FUNCTION_BLOCK Actuator2OpBaseExt (* Composite Function Block Type *)
  (* Standard: 61499-2 *)
  (* Version 1.0.1, 9/20/2023, ApplicationLibDevTeam, Schneider Electric, First Version *)
  PACKAGE Flexbridge.FestoMPS400;
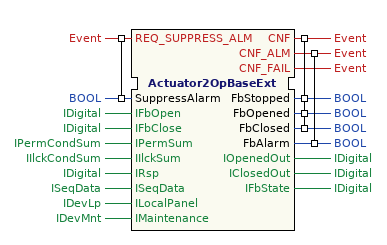
  EVENT_INPUT
    REQ_SUPPRESS_ALM WITH SuppressAlarm; (* Request to update the alarm suppress status *)
  END_EVENT
  EVENT_OUTPUT
    CNF WITH FbClosed, FbStopped, FbOpened; (* Execution confirmation *)
    CNF_ALM WITH FbAlarm; (* Execution confirmation of alarm *)
    CNF_FAIL; (* Execution confirmation of failure *)
  END_EVENT
  VAR_INPUT
    SuppressAlarm : BOOL; (* 1 = Suppress alarm in HMI *)
  END_VAR
  VAR_OUTPUT
    FbStopped : BOOL; (* 1 = Stopped *)
    FbOpened : BOOL; (* 1 = Open *)
    FbClosed : BOOL; (* 1 = Closed *)
    FbAlarm : BOOL; (* 1 = Feedback failure alarm is active *)
  END_VAR
  SOCKETS
    IFbOpen : IDigital; (* Open feedback signal adapter *)
    IFbClose : IDigital; (* Closed feedback signal adapter *)
    IPermSum : IPermCondSum(DeviceType := BiDirectional, ServiceState := TRUE); (* Permission condition summary chain input from permcondsum block *)
    IIlckSum : IIlckCondSum(DeviceType := BiDirectional, ServiceState := TRUE); (* Interlock condition summary chain input from ilckcondsum block *)
  END_SOCKETS
  SOCKETS
    IRsp : IDigital; (* Program remote setpoint interface adapter *)
    ISeqData : ISeqData; (* Sequence control interface adapter, Controls the block when owner is in program local *)
    ILocalPanel : IDevLp; (* Local panel Interface adapter *)
    IMaintenance : IDevMnt; (* Maintenance data Interface adapter *)
  END_SOCKETS
  PLUGS
    IOpenedOut : IDigital; (* Current Open Output status Interface adapter( Value = device output, Status = Bit 1 = Simulation mode) *)
    IClosedOut : IDigital; (* Current Close Output status Interface adapter( Value = device output, Status = Bit 1 = Simulation mode) *)
    IFbState : IDigital; (* Current feedback status Interface adapter(Value = device feedback status, Status = device alarm data,Bit 1 = Device failure status, Bit 2 = Feedback failure status) *)
  END_PLUGS
  (* Control *)
  (* Permissive *)
  (* Interlock *)
  (* Input Hardware Interface *)
  (* Service Connection *)
  (* Output Interface *)
  (* Hardware Output Interface *)
  FBS
    fbOpenConv : intToBool;
    invertFeedback : NOT_42C76073DCEB1A7A; {SET_ATTRIBUTE(Configuration.GenericFBType.InterfaceParams, Runtime.Standard#CNT:=1;OUT${CNT$}:BOOL)}
    serviceManager : Valve2OpServiceManager;
    orSpeed1Speed2 : OR_88A3DD8EC65DD11C; {SET_ATTRIBUTE(Configuration.GenericFBType.InterfaceParams, Runtime.Standard#CNT:=2;OUT:BOOL)}
    outConv : ANY2ANY_82AC55F556C8F3CD; {SET_ATTRIBUTE(Configuration.GenericFBType.InterfaceParams, Runtime.Standard#CNT:=2;IN${CNT$}:BOOL,BOOL;OUT${CNT$}:INT,INT)}
    actuator2OpBase : Actuator2OpBase; {SET_ATTRIBUTE(Configuration.Component.HideUnusedPorts, )}
  END_FBS
  EVENT_CONNECTIONS
    IFbOpen.REQ TO fbOpenConv.REQ1;
    actuator2OpBase.CNF_MODE TO IOpenedOut.REQ_STATUS;
    actuator2OpBase.CNF_FB_ALM TO CNF_ALM;
    actuator2OpBase.CNF_FAIL TO CNF_FAIL;
    REQ_SUPPRESS_ALM TO actuator2OpBase.REQ_SUPPRESS_ALM;
    IPermSum.PERM_IND TO actuator2OpBase.REQ_PERM;
    IIlckSum.COND_IND TO actuator2OpBase.REQ_ILCK;
    invertFeedback.CNF TO actuator2OpBase.REQ_FB;
    actuator2OpBase.CNF_FB_STS TO IFbState.REQ;
    actuator2OpBase.CNF_ALM TO IFbState.REQ_STATUS;
    IIlckSum.CHECK_SERVICE TO IIlckSum.CNF_SERVICE;
    IPermSum.CHECK_SERVICE TO IPermSum.CNF_SERVICE;
    actuator2OpBase.CNF_MODE TO IIlckSum.REQ;
    IFbClose.REQ TO fbOpenConv.REQ2;
    fbOpenConv.CNF1 TO orSpeed1Speed2.REQ;
    fbOpenConv.CNF2 TO orSpeed1Speed2.REQ;
    orSpeed1Speed2.CNF TO invertFeedback.REQ;
    actuator2OpBase.CNF_OUT TO outConv.REQ;
    outConv.CNF TO IOpenedOut.REQ;
    outConv.CNF TO IClosedOut.REQ;
    actuator2OpBase.CNF_MODE TO IClosedOut.REQ_STATUS;
    actuator2OpBase.CNF_FB_STS TO CNF;
    actuator2OpBase.CNF_OWNER TO IIlckSum.REQ_OWNER;
  END_CONNECTIONS
  DATA_CONNECTIONS
    IIlckSum.State TO actuator2OpBase.IlckCond;
    IPermSum.PermPassive TO actuator2OpBase.PermStop;
    actuator2OpBase.AlarmStatus TO IFbState.Status;
    actuator2OpBase.FbStopped TO FbStopped;
    actuator2OpBase.FbAlarm TO FbAlarm;
    SuppressAlarm TO actuator2OpBase.SuppressAlarm;
    IIlckSum.CondType TO actuator2OpBase.IlckType;
    IIlckSum.CondPos TO actuator2OpBase.IlckPos;
    invertFeedback.OUT1 TO actuator2OpBase.FbStop;
    IFbOpen.Value TO fbOpenConv.IN1;
    actuator2OpBase.FbStatus TO IFbState.Value;
    actuator2OpBase.Maintenance TO IIlckSum.Suppress;
    actuator2OpBase.Simulation TO IOpenedOut.Status;
    IFbClose.Value TO fbOpenConv.IN2;
    orSpeed1Speed2.OUT TO invertFeedback.IN1;
    fbOpenConv.OUT1 TO orSpeed1Speed2.IN1;
    fbOpenConv.OUT2 TO orSpeed1Speed2.IN2;
    fbOpenConv.OUT1 TO actuator2OpBase.FbOpen;
    actuator2OpBase.FbClosed TO FbClosed;
    actuator2OpBase.FbOpened TO FbOpened;
    fbOpenConv.OUT2 TO actuator2OpBase.FbClose;
    IPermSum.PermActive1 TO actuator2OpBase.PermOpen;
    IPermSum.PermActive2 TO actuator2OpBase.PermClose;
    actuator2OpBase.OutOpen TO outConv.IN1;
    outConv.OUT1 TO IOpenedOut.Value;
    outConv.OUT2 TO IClosedOut.Value;
    actuator2OpBase.Simulation TO IClosedOut.Status;
    actuator2OpBase.OutClose TO outConv.IN2;
    actuator2OpBase.CurrentOwner TO IIlckSum.CurrentOwner;
  END_CONNECTIONS
  ADAPTER_CONNECTIONS
    IRsp TO serviceManager.IRsp;
    IMaintenance TO serviceManager.IMaint;
    ILocalPanel TO serviceManager.28;
    ISeqData TO serviceManager.31;
    serviceManager.14 TO actuator2OpBase.230;
  END_CONNECTIONS
END_FUNCTION_BLOCK
